RoboDK station: Celula_Polimento_FANUC.rdk

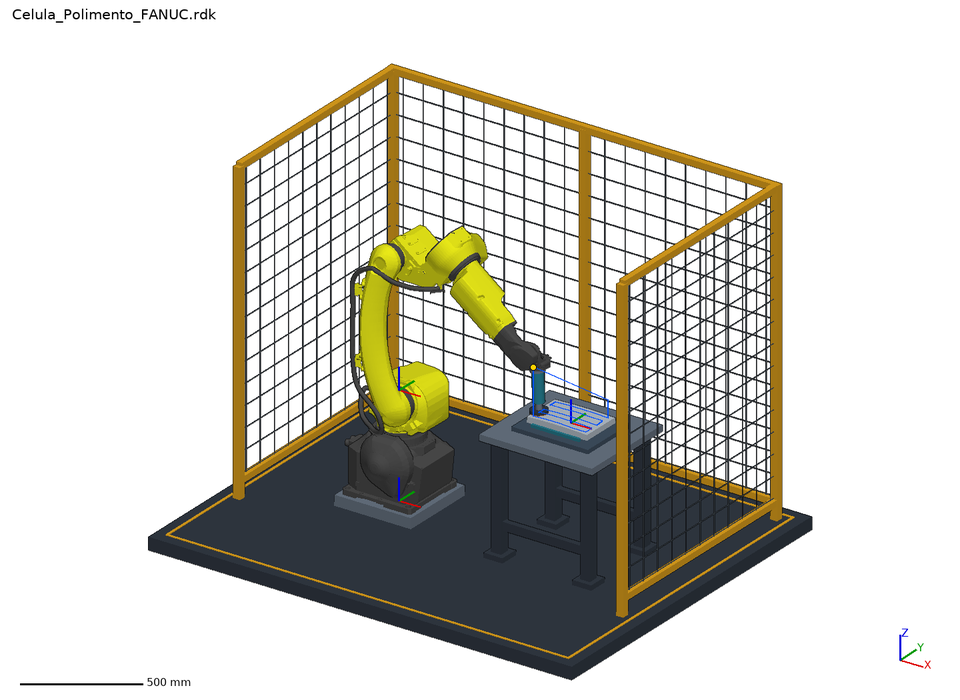
[picture v0: the station drawn from its stored meshes, robots at their saved joint values, targets as dots, program paths as lines]
Station FANUC | Polimento de tampa em aluminio (saved by RoboDK 6.0.6). Poses are relative to the parent item; angles as X-Y-Z fixed-axis rotations.
Station parameters (name, value as stored): IO_1, 1, LIN64
  - frame 01 | Estrutura da celula at (0, 0, 0) mm
    - object Plataforma at (0, 0, 0) mm, size 2100 x 1700 x 60 mm
    - object Delimitacao amarela at (0, 0, 0) mm, size 2002 x 1602 x 3 mm
    - object Placa de montagem do robo at (0, 0, 0) mm, size 380 x 380 x 50 mm
    - object Mesa - tampo at (0, 0, 0) mm, size 560 x 500 x 30 mm
    - object Mesa - estrutura at (0, 0, 0) mm, size 535 x 475 x 530 mm
    - object Base de fixacao at (0, 0, 0) mm, size 380 x 300 x 20 mm
    - object Apoios da peca at (0, 0, 0) mm, size 240 x 150 x 10 mm
    - object Batentes laterais at (0, 0, 0) mm, size 240 x 224 x 14 mm
    - object Protecao - estrutura conceptual at (0, 0, 0) mm, size 1935 x 1125 x 1515 mm
    - object Protecao - malha at (0, 0, 0) mm, size 1903 x 1091.5 x 1400 mm
  - frame 02 | Base FANUC at (0, 0, 500) mm
    - frame Fanuc M-10iD/12 Base at (0, 0, 0) mm
      - robot FANUC M-10iD/12 (model Fanuc M-10iD/12): 6 axes, payload 12 kg, reach 1441 mm, repeatability 0.02 mm, weight 145 kg
          modified DH rows (alpha deg, a mm, theta deg, d mm): 0, 0, 0, 450; -90, 75, -90, 0; 0, 640, 0, 0; -90, 195, 0, 700; 90, 0, 0, 0; -90, 0, 0, 75
          base shift (0, 0, -450) mm
          joint limits [-170, -90, -95, -190, -190, -450] to [170, 160, 180, 190, 190, 450]; home [0, 0, 0, 0, 0, 0]; saved at [-3.232, -4.4, -35.385, -0.188, -51.992, 3.344]
        - tool Polidora D80 - TCP 1, TCP at (0, 0, 200) mm, size 80 x 80 x 200 mm
  - frame 03 | Peca - UFRAME 1 at (850, 0, 590) mm
    - object Tampa aluminio 300 x 200 x 30 at (0, 0, 0) mm, size 300 x 200 x 30 mm
    - object Percurso de polimento - 5 passagens at (0, 0, 0) mm, geometry from LINEW=3
  - program POLIR (37 instructions, listed below)
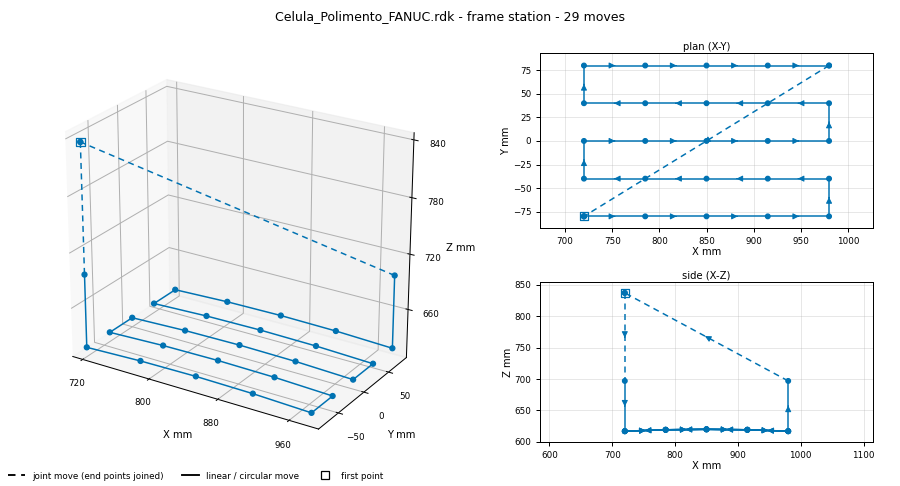
[picture p0: tool path of Celula_Polimento_FANUC.rdk in frame station, 29 of 29 moves have a stored position in this frame; points joined in program order, loops and branches not executed]

--- program POLIR (robot FANUC M-10iD/12) ---
  Set Ref.: 03 | Peca - UFRAME 1
  Set Tool: Polidora D80 - TCP 1
  Smooth(1)
  Set speed (100.0 mm/s)
  MoveJ (HOME) to (-130, -80, 247) mm, rotated rx 180 ry -2.65 rz 0 deg; joints [-6.453, -8.039, -17.302, -0.316, -70.069, 6.554]
  MoveJ (APROXIMACAO) to (-130, -80, 107) mm, rotated rx 180 ry -2.65 rz 0 deg; joints [-6.453, -6.37, -28.638, -0.348, -58.733, 6.627]
  Set IO_1=1
  Set speed (40.0 mm/s)
  MoveL (P1_1) to (-130, -80, 27) mm, rotated rx 180 ry -2.65 rz 0 deg; joints [-6.453, -4.186, -35.404, -0.377, -51.967, 6.679]
  MoveL (P1_2) to (-65, -80, 29.25) mm, rotated rx 180 ry -1.32 rz 0 deg; joints [-5.866, 2.129, -35.302, -0.169, -53.381, 5.965]
  MoveL (P1_3) to (0, -80, 30) mm, rotated rx 180 ry 0 rz 0 deg; joints [-5.377, 8.291, -34.711, 0, -55.289, 5.377]
  MoveL (P1_4) to (65, -80, 29.25) mm, rotated rx 180 ry 1.32 rz 0 deg; joints [-4.962, 14.396, -33.664, 0.136, -57.655, 4.889]
  MoveL (P1_5) to (130, -80, 27) mm, rotated rx 180 ry 2.65 rz 0 deg; joints [-4.607, 20.54, -32.168, 0.244, -60.471, 4.482]
  MoveL (P2_1) to (130, -40, 27) mm, rotated rx 180 ry 2.65 rz 0 deg; joints [-2.307, 20.333, -32.234, 0.122, -60.41, 2.245]
  MoveL (P2_2) to (65, -40, 29.25) mm, rotated rx 180 ry 1.32 rz 0 deg; joints [-2.486, 14.174, -33.715, 0.068, -57.608, 2.449]
  MoveL (P2_3) to (0, -40, 30) mm, rotated rx 180 ry 0 rz 0 deg; joints [-2.694, 8.049, -34.743, 0, -55.257, 2.694]
  MoveL (P2_4) to (-65, -40, 29.25) mm, rotated rx 180 ry -1.32 rz 0 deg; joints [-2.941, 1.857, -35.311, -0.085, -53.367, 2.99]
  MoveL (P2_5) to (-130, -40, 27) mm, rotated rx 180 ry -2.65 rz 0 deg; joints [-3.237, -4.498, -35.382, -0.19, -51.976, 3.35]
  MoveL (P3_1) to (-130, 0, 27) mm, rotated rx 180 ry -2.65 rz 0 deg; joints [0, -4.603, -35.374, 0, -51.98, 0]
  MoveL (P3_2) to (-65, 0, 29.25) mm, rotated rx 180 ry -1.32 rz 0 deg; joints [0, 1.766, -35.314, 0, -53.362, 0]
  MoveL (P3_3) to (0, 0, 30) mm, rotated rx 180 ry 0 rz 0 deg; joints [0, 7.968, -34.754, 0, -55.246, 0]
  MoveL (P3_4) to (65, 0, 29.25) mm, rotated rx 180 ry 1.32 rz 0 deg; joints [0, 14.1, -33.732, 0, -57.592, 0]
  MoveL (P3_5) to (130, 0, 27) mm, rotated rx 180 ry 2.65 rz 0 deg; joints [0, 20.263, -32.256, 0, -60.39, 0]
  MoveL (P4_1) to (130, 40, 27) mm, rotated rx 180 ry 2.65 rz 0 deg; joints [2.307, 20.333, -32.234, -0.122, -60.41, -2.245]
  MoveL (P4_2) to (65, 40, 29.25) mm, rotated rx 180 ry 1.32 rz 0 deg; joints [2.486, 14.174, -33.715, -0.068, -57.608, -2.449]
  MoveL (P4_3) to (0, 40, 30) mm, rotated rx 180 ry 0 rz 0 deg; joints [2.694, 8.049, -34.743, 0, -55.257, -2.694]
  MoveL (P4_4) to (-65, 40, 29.25) mm, rotated rx 180 ry -1.32 rz 0 deg; joints [2.941, 1.857, -35.311, 0.085, -53.367, -2.99]
  MoveL (P4_5) to (-130, 40, 27) mm, rotated rx 180 ry -2.65 rz 0 deg; joints [3.237, -4.498, -35.382, 0.19, -51.976, -3.35]
  MoveL (P5_1) to (-130, 80, 27) mm, rotated rx 180 ry -2.65 rz 0 deg; joints [6.453, -4.186, -35.404, 0.377, -51.967, -6.679]
  MoveL (P5_2) to (-65, 80, 29.25) mm, rotated rx 180 ry -1.32 rz 0 deg; joints [5.866, 2.129, -35.302, 0.169, -53.381, -5.965]
  MoveL (P5_3) to (0, 80, 30) mm, rotated rx 180 ry 0 rz 0 deg; joints [5.377, 8.291, -34.711, 0, -55.289, -5.377]
  MoveL (P5_4) to (65, 80, 29.25) mm, rotated rx 180 ry 1.32 rz 0 deg; joints [4.962, 14.396, -33.664, -0.136, -57.655, -4.889]
  MoveL (P5_5) to (130, 80, 27) mm, rotated rx 180 ry 2.65 rz 0 deg; joints [4.607, 20.54, -32.168, -0.244, -60.471, -4.482]
  MoveL (AFASTAMENTO) to (130, 80, 107) mm, rotated rx 180 ry 2.65 rz 0 deg; joints [4.607, 18.845, -26.192, -0.232, -66.446, -4.51]
  Set IO_1=0
  Set speed (100.0 mm/s)
  MoveJ (HOME) to (-130, -80, 247) mm, rotated rx 180 ry -2.65 rz 0 deg; joints [-6.453, -8.039, -17.302, -0.316, -70.069, 6.554]
